Staubli VAL3: HMI_action.pjx

--- HMI_action.pjx ---
Parameters version=s8.10.3Cs9_BS2093 stackSize=5000 millimeterUnit=true
Program file=bind.pgx
Program file=main.pgx
Program file=onSave.pgx
Program file=onShow.pgx
Program file=onStart.pgx
Program file=start.pgx
Program file=stop.pgx
Data file=HMI_action.dtx
Library alias=util path=Disk://HMI_cs9/HMI_util/HMI_util.pjx
Library alias=io path=Disk://source/projectSource/io/io.pjx
Library alias=action path=Disk://source/projectSource/Action/Action.pjx
Library alias=actdata path=Disk://data/actionData/actionData.pjx
Type name=actItem path=Disk://source/template/actItem/actItem.pjx

--- HMI_action.dtx ---
mdesc mNomSpeed
string sActionList
public string sIOList
string sSelList
string sSelIO[6]
public string sComment
bool bBack
bool bConfirm
num nSelList
string sLastList
bool bOnsave
public actItem aEditItem
  [0]
    string sComment
    actionItem aActItem[6]
      [0]
        num nIOindex
        num nboolValue
        num nPulseValue
        string sIOtype
        string sValue
        bool bActive
      [1]
        num nIOindex
        num nboolValue
        num nPulseValue
        string sIOtype
        string sValue
        bool bActive
      [2]
        num nIOindex
        num nboolValue
        num nPulseValue
        string sIOtype
        string sValue
        bool bActive
      [3]
        num nIOindex
        num nboolValue
        num nPulseValue
        string sIOtype
        string sValue
        bool bActive
      [4]
        num nIOindex
        num nboolValue
        num nPulseValue
        string sIOtype
        string sValue
        bool bActive
      [5]
        num nIOindex
        num nboolValue
        num nPulseValue
        string sIOtype
        string sValue
        bool bActive

--- main.pgx ---
public program main()
  local bool l_bExit
  local bool l_bResult
  local string l_scbx
  local string l_snmb
  local num l_i
begin
  do
    if util:sPage!="action"
      util:sPage="action"
      call onStart()
      call bind()
      userPage(util:sPage)
      delay(0.5)
    endIf
    //list
    if sSelList!=sLastList and sSelList!="--"
      sLastList=sSelList
      toNum(sSelList,nSelList,l_bResult)
      call onShow()
    endIf
    //
    for l_i = 0 to size(aEditItem.aActItem)-1
      l_scbx="cbx"+toString("",20+l_i)
      l_snmb="nmb"+toString("",l_i)
      switch aEditItem.aActItem[l_i].sIOtype
        case "PULSE"
          userPageSet("action",l_scbx,"disabled",true)
          userPageSet("action",l_snmb,"disabled",false)
        break
        case "IN","OUT"
          userPageSet("action",l_scbx,"disabled",false)
          userPageSet("action",l_snmb,"disabled",true)
        break
        default
        break
      endSwitch
    endFor
    //button
    if bBack==true
      bBack=false

      l_bExit=true
    elseIf bConfirm==true
      bConfirm=false
      call onSave()
    endIf
    delay(0)
  until l_bExit==true
end

--- start.pgx ---
program start()
begin
end

--- bind.pgx ---
public program bind()
  local string l_scbx
  local num l_i
  local string l_snum
  local string l_schk
begin
  //cbxlist
  userPageBind("action","cbxlist","options",sActionList,size(sActionList),"r")
  //cbx0
  //  for l_i = 0 to 5
  //    l_scbx="cbx"+toString("",l_i)
  //  userPageBind("action","cbx0","options",sIOList,49,"r")
  //  userPageBind("action","cbx1","options",sIOList,49,"r")
  //  userPageBind("action","cbx2","options",sIOList,49,"r")
  //  userPageBind("action","cbx3","options",sIOList,49,"r")
  //  userPageBind("action","cbx4","options",sIOList,49,"r")
  //  userPageBind("action","cbx5","options",sIOList,49,"r")
  //endFor
  //value
  userPageBind("action","cbxlist","value",sSelList,1,"rw")
  //
  for l_i = 0 to 5
    l_scbx="cbx"+toString("",l_i)
    userPageBind("action",l_scbx,"value",sSelIO[l_i],1,"rw")
    l_scbx="cbx"+toString("",10+l_i)
    userPageBind("action",l_scbx,"value",aEditItem.aActItem[l_i].sIOtype,1,"rw")
    l_scbx="cbx"+toString("",20+l_i)
    userPageBind("action",l_scbx,"value",aEditItem.aActItem[l_i].sValue,1,"rw")
  endFor
  //text
  userPageBind("action","txt1","value",aEditItem.sComment,1,"rw")
  //
  //num input
  for l_i = 0 to 5
    l_snum="nmb"+toString("",l_i)
    userPageBind("action",l_snum,"value",aEditItem.aActItem[l_i].nPulseValue,1,"rw")
  endFor

  //click
  userPageBindClick("action","btnback",bBack,true)
  userPageBindClick("action","btn1",bConfirm,true)
  //check
  for l_i = 0 to 5
    l_schk="chk"+toString("",l_i)
    userPageBind("action",l_schk,"checked",aEditItem.aActItem[l_i].bActive,1,"rw")
  endFor
end

--- onSave.pgx ---
program onSave()
  local bool l_bResult
  local num l_i
begin
  actdata:aActItem[nSelList].sComment=aEditItem.sComment
  for l_i = 0 to size(aEditItem.aActItem)-1
    actdata:aActItem[nSelList].aActItem[l_i].sIOtype=aEditItem.aActItem[l_i].sIOtype
    actdata:aActItem[nSelList].aActItem[l_i].sValue=aEditItem.aActItem[l_i].sValue
    actdata:aActItem[nSelList].aActItem[l_i].bActive=(aEditItem.aActItem[l_i].bActive==true)
    toNum(sSelIO[l_i],actdata:aActItem[nSelList].aActItem[l_i].nIOindex,l_bResult)
    if !l_bResult
      actdata:aActItem[nSelList].aActItem[l_i].nIOindex=-1
    endIf
    actdata:aActItem[nSelList].aActItem[l_i].nPulseValue=aEditItem.aActItem[l_i].nPulseValue
  endFor
  bOnsave=true
  actdata:libSave()
  delay(0.1)
end

--- onShow.pgx ---
public program onShow()
  local num l_i
begin
  aEditItem.sComment=actdata:aActItem[nSelList].sComment
  for l_i = 0 to size(aEditItem.aActItem)-1

    aEditItem.aActItem[l_i].nIOindex=actdata:aActItem[nSelList].aActItem[l_i].nIOindex
    aEditItem.aActItem[l_i].bActive=(actdata:aActItem[nSelList].aActItem[l_i].bActive==true)
    aEditItem.aActItem[l_i].nboolValue=actdata:aActItem[nSelList].aActItem[l_i].nboolValue
    aEditItem.aActItem[l_i].nPulseValue=actdata:aActItem[nSelList].aActItem[l_i].nPulseValue
    aEditItem.aActItem[l_i].sIOtype=actdata:aActItem[nSelList].aActItem[l_i].sIOtype
    aEditItem.aActItem[l_i].sValue=actdata:aActItem[nSelList].aActItem[l_i].sValue

    sSelIO[l_i]=toString("",aEditItem.aActItem[l_i].nIOindex)
  endFor
end

--- onStart.pgx ---
public program onStart()
  local num l_i
begin
  //list
  resize(sActionList,1,size(actdata:aActItem))
  for l_i = 0 to size(sActionList)-1
    sActionList[l_i]=toString("",l_i)+","+actdata:aActItem[l_i].sComment
  endFor
  //
  //  resize(sIOList,1,size(io:dInItem))
  //  for l_i = 0 to size(sIOList)-1
  //    sIOList[l_i]=toString("",l_i)
  //  endFor
  //  //
  insert(sActionList[0])
  sActionList[0]="--"
  //insert(sIOList[0])
  sLastList=""
  sSelIO="--"
end

--- stop.pgx ---
program stop()
begin
end
